FUNCTION_BLOCK basicMGEGenerico (* Logica unica do multimedidor (PM5300): valores, falta de fase, tensao e corrente H/L, comunicacao *)
  (* Standard: 61499-2 *)
  (* Version 1.5, 15/10/2026, Hidryco, Hidryco, 1.5: valores na IHM com prefixo STS_ (STS_TENSAO_AB ... STS_FREQUENCIA). 1.4: corrente A, B e C baixa (um ajuste, 3 alarmes). 1.3: so as grandezas, ajustes e alarmes da especificacao; referencia 0 = desligado; um tempo por grupo. 1.2: lista de alarmes do cliente. 1.1: frequencia como LINT (VTQLINT do PM53xxMbtcp). 1.0: PM5300 pelo HW CAT PM53xxMbtcp; falta de fase, tensao H/L e corrente H/L ajustaveis na IHM *)
  PACKAGE Hidryco.HidrycoLib;
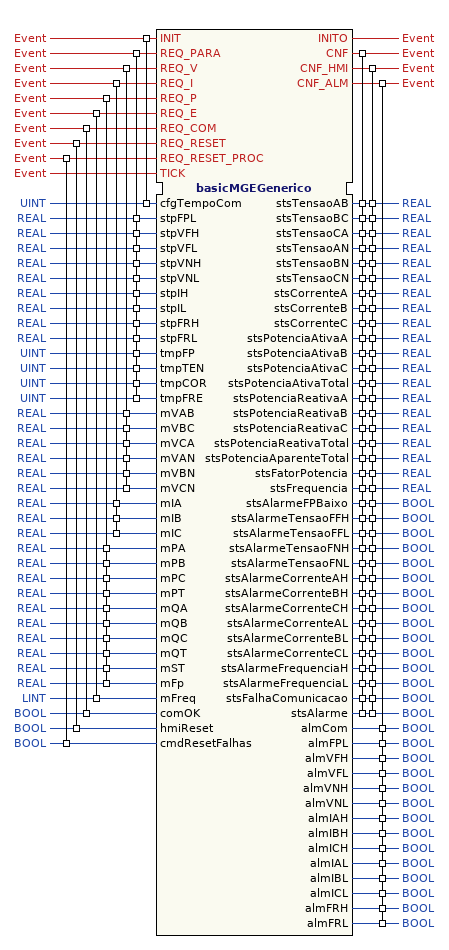
  EVENT_INPUT
    INIT WITH cfgTempoCom; (* Inicializacao *)
    REQ_PARA WITH stpFPL, stpVFH, stpVFL, stpVNH, stpVNL, stpIH, stpIL, stpFRH, stpFRL, tmpFP, tmpTEN, tmpCOR, tmpFRE; (* Parametros da IHM (persistentes) *)
    REQ_V WITH mVAB, mVBC, mVCA, mVAN, mVBN, mVCN; (* Tensoes *)
    REQ_I WITH mIA, mIB, mIC; (* Correntes *)
    REQ_P WITH mPA, mPB, mPC, mPT, mQA, mQB, mQC, mQT, mST, mFp; (* Potencias e FP *)
    REQ_E WITH mFreq; (* Frequencia *)
    REQ_COM WITH comOK; (* Comunicacao *)
    REQ_RESET WITH hmiReset; (* Reset pela IHM *)
    REQ_RESET_PROC WITH cmdResetFalhas; (* Reset pelo processo *)
    TICK; (* Base de tempo de 1 s (E_CYCLE) *)
  END_EVENT
  EVENT_OUTPUT
    INITO; (* Inicializacao concluida *)
    CNF WITH stsTensaoAB, stsTensaoBC, stsTensaoCA, stsTensaoAN, stsTensaoBN, stsTensaoCN, stsCorrenteA, stsCorrenteB, stsCorrenteC, stsPotenciaAtivaA, stsPotenciaAtivaB, stsPotenciaAtivaC, stsPotenciaAtivaTotal, stsPotenciaReativaA, stsPotenciaReativaB, stsPotenciaReativaC, stsPotenciaReativaTotal, stsPotenciaAparenteTotal, stsFatorPotencia, stsFrequencia, stsAlarmeFPBaixo, stsAlarmeTensaoFFH, stsAlarmeTensaoFFL, stsAlarmeTensaoFNH, stsAlarmeTensaoFNL, stsAlarmeCorrenteAH, stsAlarmeCorrenteBH, stsAlarmeCorrenteCH, stsAlarmeCorrenteAL, stsAlarmeCorrenteBL, stsAlarmeCorrenteCL, stsAlarmeFrequenciaH, stsAlarmeFrequenciaL, stsFalhaComunicacao, stsAlarme; (* Valores e alarmes (na mudanca) *)
    CNF_HMI WITH stsTensaoAB, stsTensaoBC, stsTensaoCA, stsTensaoAN, stsTensaoBN, stsTensaoCN, stsCorrenteA, stsCorrenteB, stsCorrenteC, stsPotenciaAtivaA, stsPotenciaAtivaB, stsPotenciaAtivaC, stsPotenciaAtivaTotal, stsPotenciaReativaA, stsPotenciaReativaB, stsPotenciaReativaC, stsPotenciaReativaTotal, stsPotenciaAparenteTotal, stsFatorPotencia, stsFrequencia, stsAlarmeFPBaixo, stsAlarmeTensaoFFH, stsAlarmeTensaoFFL, stsAlarmeTensaoFNH, stsAlarmeTensaoFNL, stsAlarmeCorrenteAH, stsAlarmeCorrenteBH, stsAlarmeCorrenteCH, stsAlarmeCorrenteAL, stsAlarmeCorrenteBL, stsAlarmeCorrenteCL, stsAlarmeFrequenciaH, stsAlarmeFrequenciaL, stsFalhaComunicacao, stsAlarme; (* Status para a IHM (na mudanca) *)
    CNF_ALM WITH almCom, almFPL, almVFH, almVFL, almVNH, almVNL, almIAH, almIBH, almICH, almIAL, almIBL, almICL, almFRH, almFRL; (* Alarmes para os ALARM_BIT (na mudanca) *)
  END_EVENT
  VAR_INPUT
    cfgTempoCom : UINT := 5; (* Tempo (s) sem comunicacao com o medidor para confirmar a falha *)
    stpFPL : REAL; (* IHM: valor de referencia - Fator de potência baixo (abaixo de) (0 = desligado) *)
    stpVFH : REAL; (* IHM: valor de referencia - Tensão entre fases alta (acima de) (0 = desligado) *)
    stpVFL : REAL; (* IHM: valor de referencia - Tensão entre fases baixa (abaixo de) (0 = desligado) *)
    stpVNH : REAL; (* IHM: valor de referencia - Tensão fase-neutro alta (acima de) (0 = desligado) *)
    stpVNL : REAL; (* IHM: valor de referencia - Tensão fase-neutro baixa (abaixo de) (0 = desligado) *)
    stpIH : REAL; (* IHM: valor de referencia - Corrente alta - fases A, B e C (acima de) (0 = desligado) *)
    stpIL : REAL; (* IHM: valor de referencia - Corrente baixa - fases A, B e C (abaixo de) (0 = desligado) *)
    stpFRH : REAL; (* IHM: valor de referencia - Frequência alta (acima de) (0 = desligado) *)
    stpFRL : REAL; (* IHM: valor de referencia - Frequência baixa (abaixo de) (0 = desligado) *)
    tmpFP : UINT; (* IHM: tempo de retardo (s) dos alarmes de fator de potência *)
    tmpTEN : UINT; (* IHM: tempo de retardo (s) dos alarmes de tensão *)
    tmpCOR : UINT; (* IHM: tempo de retardo (s) dos alarmes de corrente *)
    tmpFRE : UINT; (* IHM: tempo de retardo (s) dos alarmes de frequência *)
    mVAB : REAL; (* Tensao A-B (V) *)
    mVBC : REAL; (* Tensao B-C (V) *)
    mVCA : REAL; (* Tensao C-A (V) *)
    mVAN : REAL; (* Tensao A-N (V) *)
    mVBN : REAL; (* Tensao B-N (V) *)
    mVCN : REAL; (* Tensao C-N (V) *)
    mIA : REAL; (* Corrente fase A (A) *)
    mIB : REAL; (* Corrente fase B (A) *)
    mIC : REAL; (* Corrente fase C (A) *)
    mPA : REAL; (* Potencia ativa fase A (kW) *)
    mPB : REAL; (* Potencia ativa fase B (kW) *)
    mPC : REAL; (* Potencia ativa fase C (kW) *)
    mPT : REAL; (* Potencia ativa total (kW) *)
    mQA : REAL; (* Potencia reativa fase A (kVAr) *)
    mQB : REAL; (* Potencia reativa fase B (kVAr) *)
    mQC : REAL; (* Potencia reativa fase C (kVAr) *)
    mQT : REAL; (* Potencia reativa total (kVAr) *)
    mST : REAL; (* Potencia aparente total (kVA) *)
    mFp : REAL; (* Fator de potencia total () *)
    mFreq : LINT; (* Frequencia (Hz; o PM53xxMbtcp publica como VTQLINT, sem decimais) *)
    comOK : BOOL; (* ComStatus do PM53xxMbtcp (TRUE = comunicacao ativa) *)
    hmiReset : BOOL; (* IHM: reset / reconhecimento *)
    cmdResetFalhas : BOOL; (* Processo: reset (com E_RESET_FALHAS) *)
  END_VAR
  VAR_OUTPUT
    stsTensaoAB : REAL; (* Tensao A-B (V) *)
    stsTensaoBC : REAL; (* Tensao B-C (V) *)
    stsTensaoCA : REAL; (* Tensao C-A (V) *)
    stsTensaoAN : REAL; (* Tensao A-N (V) *)
    stsTensaoBN : REAL; (* Tensao B-N (V) *)
    stsTensaoCN : REAL; (* Tensao C-N (V) *)
    stsCorrenteA : REAL; (* Corrente fase A (A) *)
    stsCorrenteB : REAL; (* Corrente fase B (A) *)
    stsCorrenteC : REAL; (* Corrente fase C (A) *)
    stsPotenciaAtivaA : REAL; (* Potencia ativa fase A (kW) *)
    stsPotenciaAtivaB : REAL; (* Potencia ativa fase B (kW) *)
    stsPotenciaAtivaC : REAL; (* Potencia ativa fase C (kW) *)
    stsPotenciaAtivaTotal : REAL; (* Potencia ativa total (kW) *)
    stsPotenciaReativaA : REAL; (* Potencia reativa fase A (kVAr) *)
    stsPotenciaReativaB : REAL; (* Potencia reativa fase B (kVAr) *)
    stsPotenciaReativaC : REAL; (* Potencia reativa fase C (kVAr) *)
    stsPotenciaReativaTotal : REAL; (* Potencia reativa total (kVAr) *)
    stsPotenciaAparenteTotal : REAL; (* Potencia aparente total (kVA) *)
    stsFatorPotencia : REAL; (* Fator de potencia total *)
    stsFrequencia : REAL; (* Frequencia (Hz) *)
    stsAlarmeFPBaixo : BOOL; (* Fator de potência baixo (memorizado ate o reconhecimento) *)
    stsAlarmeTensaoFFH : BOOL; (* Tensão entre fases alta (memorizado ate o reconhecimento) *)
    stsAlarmeTensaoFFL : BOOL; (* Tensão entre fases baixa (memorizado ate o reconhecimento) *)
    stsAlarmeTensaoFNH : BOOL; (* Tensão fase-neutro alta (memorizado ate o reconhecimento) *)
    stsAlarmeTensaoFNL : BOOL; (* Tensão fase-neutro baixa (memorizado ate o reconhecimento) *)
    stsAlarmeCorrenteAH : BOOL; (* Corrente fase A alta (memorizado ate o reconhecimento) *)
    stsAlarmeCorrenteBH : BOOL; (* Corrente fase B alta (memorizado ate o reconhecimento) *)
    stsAlarmeCorrenteCH : BOOL; (* Corrente fase C alta (memorizado ate o reconhecimento) *)
    stsAlarmeCorrenteAL : BOOL; (* Corrente fase A baixa (memorizado ate o reconhecimento) *)
    stsAlarmeCorrenteBL : BOOL; (* Corrente fase B baixa (memorizado ate o reconhecimento) *)
    stsAlarmeCorrenteCL : BOOL; (* Corrente fase C baixa (memorizado ate o reconhecimento) *)
    stsAlarmeFrequenciaH : BOOL; (* Frequência alta (memorizado ate o reconhecimento) *)
    stsAlarmeFrequenciaL : BOOL; (* Frequência baixa (memorizado ate o reconhecimento) *)
    stsFalhaComunicacao : BOOL; (* Falha de comunicacao com o medidor *)
    stsAlarme : BOOL; (* Algum alarme do medidor *)
    almCom : BOOL; (* ALARM_BIT falha de comunicacao *)
    almFPL : BOOL; (* ALARM_BIT Fator de potência baixo *)
    almVFH : BOOL; (* ALARM_BIT Tensão entre fases alta *)
    almVFL : BOOL; (* ALARM_BIT Tensão entre fases baixa *)
    almVNH : BOOL; (* ALARM_BIT Tensão fase-neutro alta *)
    almVNL : BOOL; (* ALARM_BIT Tensão fase-neutro baixa *)
    almIAH : BOOL; (* ALARM_BIT Corrente fase A alta *)
    almIBH : BOOL; (* ALARM_BIT Corrente fase B alta *)
    almICH : BOOL; (* ALARM_BIT Corrente fase C alta *)
    almIAL : BOOL; (* ALARM_BIT Corrente fase A baixa *)
    almIBL : BOOL; (* ALARM_BIT Corrente fase B baixa *)
    almICL : BOOL; (* ALARM_BIT Corrente fase C baixa *)
    almFRH : BOOL; (* ALARM_BIT Frequência alta *)
    almFRL : BOOL; (* ALARM_BIT Frequência baixa *)
  END_VAR
  VAR
    initDone : BOOL;
    initPass : BOOL;
    bReset : BOOL;
    bComRecebida : BOOL; (* Ja houve leitura do ComStatus *)
    bValido : BOOL; (* Medidor comunicando: valores validos *)
    uSegCom : UDINT;
    cFPL : BOOL; (* Condicao agora *)
    cVFH : BOOL; (* Condicao agora *)
    cVFL : BOOL; (* Condicao agora *)
    cVNH : BOOL; (* Condicao agora *)
    cVNL : BOOL; (* Condicao agora *)
    cIAH : BOOL; (* Condicao agora *)
    cIBH : BOOL; (* Condicao agora *)
    cICH : BOOL; (* Condicao agora *)
    cIAL : BOOL; (* Condicao agora *)
    cIBL : BOOL; (* Condicao agora *)
    cICL : BOOL; (* Condicao agora *)
    cFRH : BOOL; (* Condicao agora *)
    cFRL : BOOL; (* Condicao agora *)
    uFPL : UDINT; (* Segundos na condicao *)
    uVFH : UDINT; (* Segundos na condicao *)
    uVFL : UDINT; (* Segundos na condicao *)
    uVNH : UDINT; (* Segundos na condicao *)
    uVNL : UDINT; (* Segundos na condicao *)
    uIAH : UDINT; (* Segundos na condicao *)
    uIBH : UDINT; (* Segundos na condicao *)
    uICH : UDINT; (* Segundos na condicao *)
    uIAL : UDINT; (* Segundos na condicao *)
    uIBL : UDINT; (* Segundos na condicao *)
    uICL : UDINT; (* Segundos na condicao *)
    uFRH : UDINT; (* Segundos na condicao *)
    uFRL : UDINT; (* Segundos na condicao *)
    rOld : REAL;
    bMudou : BOOL;
    wSts : WORD;
    oldSts : WORD := 16#FFFF;
    wAlm : WORD;
    oldAlm : WORD := 16#FFFF;
    o_stsTensaoAB : REAL := -1.0;
    o_stsTensaoBC : REAL := -1.0;
    o_stsTensaoCA : REAL := -1.0;
    o_stsTensaoAN : REAL := -1.0;
    o_stsTensaoBN : REAL := -1.0;
    o_stsTensaoCN : REAL := -1.0;
    o_stsCorrenteA : REAL := -1.0;
    o_stsCorrenteB : REAL := -1.0;
    o_stsCorrenteC : REAL := -1.0;
    o_stsPotenciaAtivaA : REAL := -1.0;
    o_stsPotenciaAtivaB : REAL := -1.0;
    o_stsPotenciaAtivaC : REAL := -1.0;
    o_stsPotenciaAtivaTotal : REAL := -1.0;
    o_stsPotenciaReativaA : REAL := -1.0;
    o_stsPotenciaReativaB : REAL := -1.0;
    o_stsPotenciaReativaC : REAL := -1.0;
    o_stsPotenciaReativaTotal : REAL := -1.0;
    o_stsPotenciaAparenteTotal : REAL := -1.0;
    o_stsFatorPotencia : REAL := -1.0;
    o_stsFrequencia : REAL := -1.0;
  END_VAR
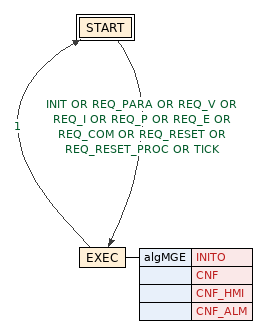
  EC_STATES
    START; (* Estado inicial *)
    EXEC : algMGE -> INITO, -> CNF, -> CNF_HMI, -> CNF_ALM; (* Executa a logica; o algoritmo decide quais eventos saem *)
  END_STATES
  EC_TRANSITIONS
    START TO EXEC := INIT OR REQ_PARA OR REQ_V OR REQ_I OR REQ_P OR REQ_E OR REQ_COM OR REQ_RESET OR REQ_RESET_PROC OR TICK;
    EXEC TO START := 1;
  END_TRANSITIONS
  ALGORITHM algMGE IN ST: (* Logica completa do multimedidor (um unico algoritmo) *)
(* =====================================================================
   basicMGEGenerico v1.5 - multimedidor PowerLogic PM5300 (HW CAT PM53xxMbtcp)
   Padrao das bibliotecas Schneider: eventos de saida desligados no inicio e
   ligados so na mudanca; tempos contados pelo TICK de 1 s (E_CYCLE do CAT).
   - valores recebidos dos symlinks VTQ do PM53xxMbtcp; energias de Wh para kWh;
   - v1.1: frequencia recebida como VTQLINT (e assim que o PM53xxMbtcp publica);
   - falha de comunicacao: ComStatus FALSE por cfgTempoCom s; com a falha,
     os alarmes de medicao ficam suprimidos (os valores ficam congelados);
   - v1.2: falta de fase (FF abaixo do ajuste); tensao entre fases e
     fase-neutro alta/baixa (as baixas nao atuam junto com a falta de
     fase); corrente A, B e C alta (um ajuste, 3 alarmes); FP baixo (so
     com carga: potencia aparente > 0); frequencia alta/baixa;
   - v1.3: so as grandezas e alarmes da especificacao (sai a falta de fase,
     as medias, o desequilibrio, a aparente por fase e as energias); valor
     de referencia por limite (0 = desligado) e um tempo de retardo por
     grupo (FP, tensao, corrente, frequencia); memorizado ate o
     reconhecimento, que so libera o que ja normalizou;
   - v1.4: corrente A, B e C baixa (um ajuste, 3 alarmes, retardo do
     grupo corrente).
   ===================================================================== *)

INITO   := FALSE;
CNF     := FALSE;
CNF_HMI := FALSE;
CNF_ALM := FALSE;

IF REQ_COM THEN
    bComRecebida := TRUE;
END_IF;
IF INIT THEN
    initDone := TRUE;
    initPass := TRUE;
    INITO    := TRUE;
END_IF;
IF NOT initDone THEN
    RETURN;
END_IF;
bReset := (REQ_RESET AND hmiReset) OR (REQ_RESET_PROC AND cmdResetFalhas);

(* ---- 1. Comunicacao ---- *)
IF NOT comOK THEN
    IF TICK AND uSegCom < UINT_TO_UDINT(cfgTempoCom) THEN
        uSegCom := uSegCom + 1;
    END_IF;
ELSE
    uSegCom := 0;
END_IF;
stsFalhaComunicacao := NOT comOK AND uSegCom >= UINT_TO_UDINT(cfgTempoCom);
bValido := bComRecebida AND comOK;

(* ---- 2. Valores ---- *)
stsTensaoAB := mVAB;
stsTensaoBC := mVBC;
stsTensaoCA := mVCA;
stsTensaoAN := mVAN;
stsTensaoBN := mVBN;
stsTensaoCN := mVCN;
stsCorrenteA := mIA;
stsCorrenteB := mIB;
stsCorrenteC := mIC;
stsPotenciaAtivaA := mPA;
stsPotenciaAtivaB := mPB;
stsPotenciaAtivaC := mPC;
stsPotenciaAtivaTotal := mPT;
stsPotenciaReativaA := mQA;
stsPotenciaReativaB := mQB;
stsPotenciaReativaC := mQC;
stsPotenciaReativaTotal := mQT;
stsPotenciaAparenteTotal := mST;
stsFatorPotencia := mFp;
stsFrequencia := LINT_TO_REAL(mFreq);

(* ---- 3. Condicoes (so com o medidor comunicando) ---- *)
cFPL := stpFPL > 0.0 AND bValido AND (mST > 0.0 AND ABS(mFp) < stpFPL);
cVFH := stpVFH > 0.0 AND bValido AND (mVAB > stpVFH OR mVBC > stpVFH OR mVCA > stpVFH);
cVFL := stpVFL > 0.0 AND bValido AND (mVAB < stpVFL OR mVBC < stpVFL OR mVCA < stpVFL);
cVNH := stpVNH > 0.0 AND bValido AND (mVAN > stpVNH OR mVBN > stpVNH OR mVCN > stpVNH);
cVNL := stpVNL > 0.0 AND bValido AND (mVAN < stpVNL OR mVBN < stpVNL OR mVCN < stpVNL);
cIAH := stpIH > 0.0 AND bValido AND (mIA > stpIH);
cIBH := stpIH > 0.0 AND bValido AND (mIB > stpIH);
cICH := stpIH > 0.0 AND bValido AND (mIC > stpIH);
cIAL := stpIL > 0.0 AND bValido AND (mIA < stpIL);
cIBL := stpIL > 0.0 AND bValido AND (mIB < stpIL);
cICL := stpIL > 0.0 AND bValido AND (mIC < stpIL);
cFRH := stpFRH > 0.0 AND bValido AND (stsFrequencia > stpFRH);
cFRL := stpFRL > 0.0 AND bValido AND (stsFrequencia < stpFRL);

(* ---- 4. Alarmes: tempo de retardo do grupo, memoria ate o reset, referencia 0 zera ---- *)
IF cFPL THEN
    IF TICK AND uFPL < UINT_TO_UDINT(tmpFP) THEN
        uFPL := uFPL + 1;
    END_IF;
    IF uFPL >= UINT_TO_UDINT(tmpFP) THEN
        stsAlarmeFPBaixo := TRUE;
    END_IF;
ELSE
    uFPL := 0;
    IF bReset THEN
        stsAlarmeFPBaixo := FALSE;
    END_IF;
END_IF;
IF stpFPL <= 0.0 THEN
    stsAlarmeFPBaixo := FALSE;
END_IF;
IF cVFH THEN
    IF TICK AND uVFH < UINT_TO_UDINT(tmpTEN) THEN
        uVFH := uVFH + 1;
    END_IF;
    IF uVFH >= UINT_TO_UDINT(tmpTEN) THEN
        stsAlarmeTensaoFFH := TRUE;
    END_IF;
ELSE
    uVFH := 0;
    IF bReset THEN
        stsAlarmeTensaoFFH := FALSE;
    END_IF;
END_IF;
IF stpVFH <= 0.0 THEN
    stsAlarmeTensaoFFH := FALSE;
END_IF;
IF cVFL THEN
    IF TICK AND uVFL < UINT_TO_UDINT(tmpTEN) THEN
        uVFL := uVFL + 1;
    END_IF;
    IF uVFL >= UINT_TO_UDINT(tmpTEN) THEN
        stsAlarmeTensaoFFL := TRUE;
    END_IF;
ELSE
    uVFL := 0;
    IF bReset THEN
        stsAlarmeTensaoFFL := FALSE;
    END_IF;
END_IF;
IF stpVFL <= 0.0 THEN
    stsAlarmeTensaoFFL := FALSE;
END_IF;
IF cVNH THEN
    IF TICK AND uVNH < UINT_TO_UDINT(tmpTEN) THEN
        uVNH := uVNH + 1;
    END_IF;
    IF uVNH >= UINT_TO_UDINT(tmpTEN) THEN
        stsAlarmeTensaoFNH := TRUE;
    END_IF;
ELSE
    uVNH := 0;
    IF bReset THEN
        stsAlarmeTensaoFNH := FALSE;
    END_IF;
END_IF;
IF stpVNH <= 0.0 THEN
    stsAlarmeTensaoFNH := FALSE;
END_IF;
IF cVNL THEN
    IF TICK AND uVNL < UINT_TO_UDINT(tmpTEN) THEN
        uVNL := uVNL + 1;
    END_IF;
    IF uVNL >= UINT_TO_UDINT(tmpTEN) THEN
        stsAlarmeTensaoFNL := TRUE;
    END_IF;
ELSE
    uVNL := 0;
    IF bReset THEN
        stsAlarmeTensaoFNL := FALSE;
    END_IF;
END_IF;
IF stpVNL <= 0.0 THEN
    stsAlarmeTensaoFNL := FALSE;
END_IF;
IF cIAH THEN
    IF TICK AND uIAH < UINT_TO_UDINT(tmpCOR) THEN
        uIAH := uIAH + 1;
    END_IF;
    IF uIAH >= UINT_TO_UDINT(tmpCOR) THEN
        stsAlarmeCorrenteAH := TRUE;
    END_IF;
ELSE
    uIAH := 0;
    IF bReset THEN
        stsAlarmeCorrenteAH := FALSE;
    END_IF;
END_IF;
IF stpIH <= 0.0 THEN
    stsAlarmeCorrenteAH := FALSE;
END_IF;
IF cIBH THEN
    IF TICK AND uIBH < UINT_TO_UDINT(tmpCOR) THEN
        uIBH := uIBH + 1;
    END_IF;
    IF uIBH >= UINT_TO_UDINT(tmpCOR) THEN
        stsAlarmeCorrenteBH := TRUE;
    END_IF;
ELSE
    uIBH := 0;
    IF bReset THEN
        stsAlarmeCorrenteBH := FALSE;
    END_IF;
END_IF;
IF stpIH <= 0.0 THEN
    stsAlarmeCorrenteBH := FALSE;
END_IF;
IF cICH THEN
    IF TICK AND uICH < UINT_TO_UDINT(tmpCOR) THEN
        uICH := uICH + 1;
    END_IF;
    IF uICH >= UINT_TO_UDINT(tmpCOR) THEN
        stsAlarmeCorrenteCH := TRUE;
    END_IF;
ELSE
    uICH := 0;
    IF bReset THEN
        stsAlarmeCorrenteCH := FALSE;
    END_IF;
END_IF;
IF stpIH <= 0.0 THEN
    stsAlarmeCorrenteCH := FALSE;
END_IF;
IF cIAL THEN
    IF TICK AND uIAL < UINT_TO_UDINT(tmpCOR) THEN
        uIAL := uIAL + 1;
    END_IF;
    IF uIAL >= UINT_TO_UDINT(tmpCOR) THEN
        stsAlarmeCorrenteAL := TRUE;
    END_IF;
ELSE
    uIAL := 0;
    IF bReset THEN
        stsAlarmeCorrenteAL := FALSE;
    END_IF;
END_IF;
IF stpIL <= 0.0 THEN
    stsAlarmeCorrenteAL := FALSE;
END_IF;
IF cIBL THEN
    IF TICK AND uIBL < UINT_TO_UDINT(tmpCOR) THEN
        uIBL := uIBL + 1;
    END_IF;
    IF uIBL >= UINT_TO_UDINT(tmpCOR) THEN
        stsAlarmeCorrenteBL := TRUE;
    END_IF;
ELSE
    uIBL := 0;
    IF bReset THEN
        stsAlarmeCorrenteBL := FALSE;
    END_IF;
END_IF;
IF stpIL <= 0.0 THEN
    stsAlarmeCorrenteBL := FALSE;
END_IF;
IF cICL THEN
    IF TICK AND uICL < UINT_TO_UDINT(tmpCOR) THEN
        uICL := uICL + 1;
    END_IF;
    IF uICL >= UINT_TO_UDINT(tmpCOR) THEN
        stsAlarmeCorrenteCL := TRUE;
    END_IF;
ELSE
    uICL := 0;
    IF bReset THEN
        stsAlarmeCorrenteCL := FALSE;
    END_IF;
END_IF;
IF stpIL <= 0.0 THEN
    stsAlarmeCorrenteCL := FALSE;
END_IF;
IF cFRH THEN
    IF TICK AND uFRH < UINT_TO_UDINT(tmpFRE) THEN
        uFRH := uFRH + 1;
    END_IF;
    IF uFRH >= UINT_TO_UDINT(tmpFRE) THEN
        stsAlarmeFrequenciaH := TRUE;
    END_IF;
ELSE
    uFRH := 0;
    IF bReset THEN
        stsAlarmeFrequenciaH := FALSE;
    END_IF;
END_IF;
IF stpFRH <= 0.0 THEN
    stsAlarmeFrequenciaH := FALSE;
END_IF;
IF cFRL THEN
    IF TICK AND uFRL < UINT_TO_UDINT(tmpFRE) THEN
        uFRL := uFRL + 1;
    END_IF;
    IF uFRL >= UINT_TO_UDINT(tmpFRE) THEN
        stsAlarmeFrequenciaL := TRUE;
    END_IF;
ELSE
    uFRL := 0;
    IF bReset THEN
        stsAlarmeFrequenciaL := FALSE;
    END_IF;
END_IF;
IF stpFRL <= 0.0 THEN
    stsAlarmeFrequenciaL := FALSE;
END_IF;

almCom := stsFalhaComunicacao;
almFPL := stsAlarmeFPBaixo;
almVFH := stsAlarmeTensaoFFH;
almVFL := stsAlarmeTensaoFFL;
almVNH := stsAlarmeTensaoFNH;
almVNL := stsAlarmeTensaoFNL;
almIAH := stsAlarmeCorrenteAH;
almIBH := stsAlarmeCorrenteBH;
almICH := stsAlarmeCorrenteCH;
almIAL := stsAlarmeCorrenteAL;
almIBL := stsAlarmeCorrenteBL;
almICL := stsAlarmeCorrenteCL;
almFRH := stsAlarmeFrequenciaH;
almFRL := stsAlarmeFrequenciaL;
stsAlarme := almCom OR almFPL OR almVFH OR almVFL OR almVNH OR almVNL OR almIAH OR almIBH OR almICH OR almIAL OR almIBL OR almICL OR almFRH OR almFRL;

(* ---- 5. Eventos so na mudanca ---- *)
bMudou := FALSE;
IF stsTensaoAB <> o_stsTensaoAB THEN bMudou := TRUE; o_stsTensaoAB := stsTensaoAB; END_IF;
IF stsTensaoBC <> o_stsTensaoBC THEN bMudou := TRUE; o_stsTensaoBC := stsTensaoBC; END_IF;
IF stsTensaoCA <> o_stsTensaoCA THEN bMudou := TRUE; o_stsTensaoCA := stsTensaoCA; END_IF;
IF stsTensaoAN <> o_stsTensaoAN THEN bMudou := TRUE; o_stsTensaoAN := stsTensaoAN; END_IF;
IF stsTensaoBN <> o_stsTensaoBN THEN bMudou := TRUE; o_stsTensaoBN := stsTensaoBN; END_IF;
IF stsTensaoCN <> o_stsTensaoCN THEN bMudou := TRUE; o_stsTensaoCN := stsTensaoCN; END_IF;
IF stsCorrenteA <> o_stsCorrenteA THEN bMudou := TRUE; o_stsCorrenteA := stsCorrenteA; END_IF;
IF stsCorrenteB <> o_stsCorrenteB THEN bMudou := TRUE; o_stsCorrenteB := stsCorrenteB; END_IF;
IF stsCorrenteC <> o_stsCorrenteC THEN bMudou := TRUE; o_stsCorrenteC := stsCorrenteC; END_IF;
IF stsPotenciaAtivaA <> o_stsPotenciaAtivaA THEN bMudou := TRUE; o_stsPotenciaAtivaA := stsPotenciaAtivaA; END_IF;
IF stsPotenciaAtivaB <> o_stsPotenciaAtivaB THEN bMudou := TRUE; o_stsPotenciaAtivaB := stsPotenciaAtivaB; END_IF;
IF stsPotenciaAtivaC <> o_stsPotenciaAtivaC THEN bMudou := TRUE; o_stsPotenciaAtivaC := stsPotenciaAtivaC; END_IF;
IF stsPotenciaAtivaTotal <> o_stsPotenciaAtivaTotal THEN bMudou := TRUE; o_stsPotenciaAtivaTotal := stsPotenciaAtivaTotal; END_IF;
IF stsPotenciaReativaA <> o_stsPotenciaReativaA THEN bMudou := TRUE; o_stsPotenciaReativaA := stsPotenciaReativaA; END_IF;
IF stsPotenciaReativaB <> o_stsPotenciaReativaB THEN bMudou := TRUE; o_stsPotenciaReativaB := stsPotenciaReativaB; END_IF;
IF stsPotenciaReativaC <> o_stsPotenciaReativaC THEN bMudou := TRUE; o_stsPotenciaReativaC := stsPotenciaReativaC; END_IF;
IF stsPotenciaReativaTotal <> o_stsPotenciaReativaTotal THEN bMudou := TRUE; o_stsPotenciaReativaTotal := stsPotenciaReativaTotal; END_IF;
IF stsPotenciaAparenteTotal <> o_stsPotenciaAparenteTotal THEN bMudou := TRUE; o_stsPotenciaAparenteTotal := stsPotenciaAparenteTotal; END_IF;
IF stsFatorPotencia <> o_stsFatorPotencia THEN bMudou := TRUE; o_stsFatorPotencia := stsFatorPotencia; END_IF;
IF stsFrequencia <> o_stsFrequencia THEN bMudou := TRUE; o_stsFrequencia := stsFrequencia; END_IF;
wSts := 0;
IF stsAlarmeFPBaixo THEN wSts := wSts OR 16#0001; END_IF;
IF stsAlarmeTensaoFFH THEN wSts := wSts OR 16#0002; END_IF;
IF stsAlarmeTensaoFFL THEN wSts := wSts OR 16#0004; END_IF;
IF stsAlarmeTensaoFNH THEN wSts := wSts OR 16#0008; END_IF;
IF stsAlarmeTensaoFNL THEN wSts := wSts OR 16#0010; END_IF;
IF stsAlarmeCorrenteAH THEN wSts := wSts OR 16#0020; END_IF;
IF stsAlarmeCorrenteBH THEN wSts := wSts OR 16#0040; END_IF;
IF stsAlarmeCorrenteCH THEN wSts := wSts OR 16#0080; END_IF;
IF stsAlarmeCorrenteAL THEN wSts := wSts OR 16#0100; END_IF;
IF stsAlarmeCorrenteBL THEN wSts := wSts OR 16#0200; END_IF;
IF stsAlarmeCorrenteCL THEN wSts := wSts OR 16#0400; END_IF;
IF stsAlarmeFrequenciaH THEN wSts := wSts OR 16#0800; END_IF;
IF stsAlarmeFrequenciaL THEN wSts := wSts OR 16#1000; END_IF;
IF stsFalhaComunicacao THEN wSts := wSts OR 16#2000; END_IF;
IF stsAlarme THEN wSts := wSts OR 16#4000; END_IF;
wAlm := 0;
IF almCom THEN wAlm := wAlm OR 16#0001; END_IF;
IF almFPL THEN wAlm := wAlm OR 16#0002; END_IF;
IF almVFH THEN wAlm := wAlm OR 16#0004; END_IF;
IF almVFL THEN wAlm := wAlm OR 16#0008; END_IF;
IF almVNH THEN wAlm := wAlm OR 16#0010; END_IF;
IF almVNL THEN wAlm := wAlm OR 16#0020; END_IF;
IF almIAH THEN wAlm := wAlm OR 16#0040; END_IF;
IF almIBH THEN wAlm := wAlm OR 16#0080; END_IF;
IF almICH THEN wAlm := wAlm OR 16#0100; END_IF;
IF almIAL THEN wAlm := wAlm OR 16#0200; END_IF;
IF almIBL THEN wAlm := wAlm OR 16#0400; END_IF;
IF almICL THEN wAlm := wAlm OR 16#0800; END_IF;
IF almFRH THEN wAlm := wAlm OR 16#1000; END_IF;
IF almFRL THEN wAlm := wAlm OR 16#2000; END_IF;
CNF := initPass OR bMudou OR (wSts <> oldSts);
CNF_HMI := CNF;
CNF_ALM := initPass OR (wAlm <> oldAlm);
oldSts := wSts;
oldAlm := wAlm;
initPass := FALSE;
  END_ALGORITHM
END_FUNCTION_BLOCK
